Universal Robots URScript: T001_mock-model-v1_edit_lazy_rep1.urscript

def task():
  set_tcp(p[0, 0, 0.150, 0, 0, 0])
  set_payload(0.5, [0, 0, 0.05])
  movej([0, -1.57, 1.57, -1.57, -1.57, 0])
  movel(p[0.3, 0.2, 0.4, 0, 3.14, 0])
end
